(* IEC 61131-3 sources: SemaPLC/sema-plc-benchmark/spec2control-benchmark/data/st-baseline/lng-production/pous/programs, 7 files *)

(* ---- main.st ---- *)
PROGRAM main
VAR
	Heartbeat : bool;
END_VAR

(* Entry point required by OpenPLC Editor v4. The process sections run as parallel program instances under task0; main only provides a scan heartbeat. *)
Heartbeat := NOT Heartbeat;

END_PROGRAM

(* ---- Section2.st ---- *)
PROGRAM Section2
VAR
	FT_101_Flow_PV : real;
	IT_102_Flow_PV : real;
	DP_101_DiffP_PV : real;
	DP_102_DiffP_PV : real;
	LT_101_Level_PV : real;
	IIC_101_LiqSepFlow_SP : real;
	DP_101 : ANALOG_IN;
	DP_102 : ANALOG_IN;
	FT_101 : ANALOG_IN;
	IT_102 : ANALOG_IN;
	LT_101 : ANALOG_IN;
	IIC_101 : RATIO_CONTROL;
	LCV_101 : VALVE_ELECTRIC;
	LCV101_Inhibit_OR : bool;
	IIC101_Inhibit_OR : bool;
END_VAR

DP_101(
    Alarm_Enable := TRUE);
DP_102(
    Alarm_Enable := TRUE);
FT_101(
    Scaling_Slope := 312.5,
    Scaling_Offset := -1250.0,
    Alarm_Enable := TRUE);
IT_102(
    Scaling_Slope := 125.0,
    Scaling_Offset := -500.0,
    Alarm_Enable := TRUE);
LT_101(
    Alarm_Enable := TRUE);
IIC101_Inhibit_OR := LT_101.High_Alarm OR FT_101.Low_Alarm OR DP_101.High_Alarm OR DP_102.High_Alarm;
IIC_101(
    Auto := TRUE,
    PrimaryPV := FT_101.PV,
    SecondaryPV := IT_102.PV,
    RatioSP := 2.5,
    Bias := 0.0,
    MV_MIN := 0.0,
    MV_MAX := 100.0,
    Inhibit := IIC101_Inhibit_OR);
LCV101_Inhibit_OR := FT_101.Low_Alarm OR IT_102.High_Alarm OR IT_102.Low_Alarm OR DP_101.High_Alarm OR DP_102.High_Alarm;
LCV_101(
    Control_Signal := IIC_101.SlaveSP,
    Manual_Mode := FALSE,
    Open_Limit := 100.0,
    Close_Limit := 0.0,
    Inhibit := LCV101_Inhibit_OR);

(* Outputs published to other sections / HMI. *)
FT_101_Flow_PV := FT_101.PV;
IT_102_Flow_PV := IT_102.PV;
DP_101_DiffP_PV := DP_101.PV;
DP_102_DiffP_PV := DP_102.PV;
LT_101_Level_PV := LT_101.PV;
IIC_101_LiqSepFlow_SP := IIC_101.SlaveSP;

END_PROGRAM

(* ---- Section3.st ---- *)
PROGRAM Section3
VAR
	TT201_Temperature_PV : real;
	PT201_FlashTankPressure_PV : real;
	LT201_AbsorberLevel_PV : real;
	AI201_CO2_PV : real;
	TIC201_MV_SteamValveCmd : real;
	AI_201 : ANALOG_IN;
	LT_201 : ANALOG_IN;
	PT_201 : ANALOG_IN;
	TT_201 : ANALOG_IN;
	TIC_201 : PID_BASIC;
	FV_101 : VALVE_ELECTRIC;
	TIC201_Inhibit_OR : bool;
	FV101_Inhibit_OR : bool;
END_VAR

AI_201(
    Alarm_Enable := TRUE);
LT_201(
    Alarm_Enable := TRUE);
PT_201(
    PV_Low := 0.5,
    Alarm_Enable := TRUE);
TT_201(
    PV_High := 50.0,
    Scaling_Slope := 6.25,
    Scaling_Offset := -25.0,
    Alarm_Enable := TRUE);
TIC201_Inhibit_OR := TT_201.High_Alarm OR PT_201.Low_Alarm OR AI_201.High_Alarm OR TT_201.General_Fault;
FV101_Inhibit_OR := TIC201_Inhibit_OR OR LT_201.Low_Alarm;
FV_101(
    Control_Signal := TIC_201.XOUT,
    Manual_Mode := FALSE,
    Open_Limit := 100.0,
    Close_Limit := 0.0,
    Inhibit := FV101_Inhibit_OR);
TIC_201(
    AUTO := TRUE,
    PV := TT_201.PV,
    SP := 45.0,
    MV_MIN := 0.0,
    MV_MAX := 100.0,
    X0 := FV_101.Feedback_Pos,
    KP := 3.0,
    TR := 1.5,
    TD := 0.0,
    Deviation_Limit := 5.0,
    Inhibit := TIC201_Inhibit_OR);

(* Outputs published to other sections / HMI. *)
TT201_Temperature_PV := TT_201.PV;
PT201_FlashTankPressure_PV := PT_201.PV;
LT201_AbsorberLevel_PV := LT_201.PV;
AI201_CO2_PV := AI_201.PV;
TIC201_MV_SteamValveCmd := TIC_201.XOUT;

END_PROGRAM

(* ---- Section4.st ---- *)
PROGRAM Section4
VAR
	AI302_H2O_Outlet_PV : real;
	AI303_Hg_Permissive_PV : real;
	AI304_H2O_RatioOpt_PV : real;
	FT301_FeedGasFlow_PV : real;
	DP301_MolSieveBed_DP_PV : real;
	FFIC303_RegenFlow_SP_to_FIC302 : real;
	AI_302 : ANALOG_IN;
	AI_303 : ANALOG_IN;
	AI_304 : ANALOG_IN;
	DI_301 : DIGITAL_IN;
	DP_301 : ANALOG_IN;
	FIC_302 : PID_BASIC;
	FT_301 : ANALOG_IN;
	FV_302 : VALVE_ELECTRIC;
	FFIC_303 : RATIO_CONTROL;
	Inhibit_OR : bool;
END_VAR

AI_302(
    Alarm_Enable := TRUE);
AI_303(
    Alarm_Enable := TRUE);
AI_304(
    PV_High := 10.0,
    Alarm_Enable := TRUE);
DI_301();
DP_301(
    PV_High := 20.0,
    Alarm_Enable := TRUE);
FT_301(
    PV_Low := 500.0,
    Scaling_Slope := 6.25,
    Scaling_Offset := -25.0,
    Alarm_Enable := TRUE);
Inhibit_OR := AI_302.High_Alarm OR AI_303.High_Alarm OR AI_302.General_Fault OR AI_303.General_Fault OR DI_301.DI_Out OR FT_301.Low_Alarm OR DP_301.High_Alarm;
FFIC_303(
    Auto := TRUE,
    PrimaryPV := FT_301.PV,
    RatioSP := 0.25,
    Bias := 0.0,
    MV_MIN := 0.0,
    MV_MAX := 100.0,
    Inhibit := Inhibit_OR);
FIC_302(
    AUTO := TRUE,
    SP := FFIC_303.SlaveSP,
    MV_MIN := 0.0,
    MV_MAX := 100.0,
    Inhibit := Inhibit_OR);
FV_302(
    Control_Signal := FIC_302.XOUT,
    Open_Limit := 100.0,
    Close_Limit := 0.0,
    Inhibit := Inhibit_OR);

(* Outputs published to other sections / HMI. *)
AI302_H2O_Outlet_PV := AI_302.PV;
AI303_Hg_Permissive_PV := AI_303.PV;
AI304_H2O_RatioOpt_PV := AI_304.PV;
FT301_FeedGasFlow_PV := FT_301.PV;
DP301_MolSieveBed_DP_PV := DP_301.PV;
FFIC303_RegenFlow_SP_to_FIC302 := FFIC_303.SlaveSP;

END_PROGRAM

(* ---- Section5.st ---- *)
PROGRAM Section5
VAR
	PVT_401_Voted_Pressure : real;
	TVT_402_Voted_Temperature : real;
	PT_401A : ANALOG_IN;
	PT_401B : ANALOG_IN;
	PT_401C : ANALOG_IN;
	TT_105 : ANALOG_IN;
	TT_106 : ANALOG_IN;
	TT_107 : ANALOG_IN;
	PVT_401 : VOTING_ANALOG;
	TVT_402 : VOTING_ANALOG;
	PIC_401 : PID_BASIC;
	TIC_402 : PID_BASIC;
	PV_102 : VALVE_ELECTRIC;
	FV_107 : VALVE_ELECTRIC;
	XV_104 : VALVE_ON_OFF;
	I_401 : BOOL_INPUT;
	I_402 : BOOL_INPUT;
	MA_401 : BOOL_INPUT;
	PV102_Inhibit_OR : bool;
	AllPTBad_AND : bool;
	FV107_Inhibit_OR : bool;
	MasterAlarm_OR : bool;
END_VAR

PT_401A(
    PV_High := 2.0,
    PV_Low := 1.6,
    Alarm_Enable := TRUE);
PT_401B(
    PV_High := 2.0,
    PV_Low := 1.6,
    Alarm_Enable := TRUE);
PT_401C(
    PV_High := 2.0,
    PV_Low := 1.6,
    Alarm_Enable := TRUE);
TT_105(
    Alarm_Enable := TRUE);
TT_106(
    Alarm_Enable := TRUE);
TT_107(
    Alarm_Enable := TRUE);
PVT_401(
    Input1 := PT_401A.PV,
    Input2 := PT_401B.PV,
    Input3 := PT_401C.PV,
    Deviation_Limit := 0.09,
    Voting_Scheme := '2oo3',
    EnableAlarm := TRUE);
TVT_402(
    Input1 := TT_105.PV,
    Input2 := TT_106.PV,
    Input3 := TT_107.PV,
    Deviation_Limit := 2.0,
    Voting_Scheme := 'Median',
    EnableAlarm := TRUE);
PIC_401(
    AUTO := TRUE,
    PV := PVT_401.Voted_Output,
    SP := 1.8,
    MV_MIN := 0.0,
    MV_MAX := 100.0);
TIC_402(
    AUTO := TRUE,
    PV := TVT_402.Voted_Output,
    SP := 65.0,
    MV_MIN := 0.0,
    MV_MAX := 100.0);
PV102_Inhibit_OR := PVT_401.Alarm_Voting_Error OR PIC_401.PV_High_Alarm OR PIC_401.PV_Low_Alarm;
I_401(
    Bool_In := PV102_Inhibit_OR,
    Alarm_OnTrue := TRUE,
    Latch_Enable := TRUE);
PV_102(
    Control_Signal := PIC_401.XOUT,
    Open_Limit := 100.0,
    Close_Limit := 0.0,
    Timeout := T#10s,
    Inhibit := I_401.Bool_Out);
FV107_Inhibit_OR := TVT_402.Alarm_Voting_Error OR TIC_402.PV_High_Alarm OR TIC_402.PV_Low_Alarm;
I_402(
    Bool_In := FV107_Inhibit_OR,
    Alarm_OnTrue := TRUE,
    Latch_Enable := TRUE);
FV_107(
    Control_Signal := TIC_402.XOUT,
    Open_Limit := 100.0,
    Close_Limit := 0.0,
    Timeout := T#10s,
    Inhibit := I_402.Bool_Out);
AllPTBad_AND := PT_401A.General_Fault AND PT_401B.General_Fault AND PT_401C.General_Fault;
XV_104(
    Open_Cmd := FALSE,
    Close_Cmd := AllPTBad_AND,
    Timeout := T#5s,
    Inhibit := AllPTBad_AND);
MasterAlarm_OR := PV102_Inhibit_OR OR FV107_Inhibit_OR OR PT_401A.General_Fault OR PT_401B.General_Fault OR PT_401C.General_Fault OR TT_105.General_Fault OR TT_106.General_Fault OR TT_107.General_Fault;
MA_401(
    Bool_In := MasterAlarm_OR,
    Alarm_OnTrue := TRUE,
    Latch_Enable := TRUE);

(* Outputs published to other sections / HMI. *)
PVT_401_Voted_Pressure := PVT_401.Voted_Output;
TVT_402_Voted_Temperature := TVT_402.Voted_Output;

END_PROGRAM

(* ---- Section6.st ---- *)
PROGRAM Section6
VAR
	FT501_PropaneFlow_PV : real;
	FT502_MRFlow_PV : real;
	PT501_EndFlashDrumPressure_PV : real;
	TIT102_MCHE_OutletTemp_PV : real;
	FIC504_MRFlow_SP_From_FFIC503 : real;
	FFIC503_ActiveRatio : real;
	Operator_RatioBias : real;
	FFIC503_DV_HI : bool;
	FFIC503_DV_LO : bool;
	FFIC_503 : RATIO_CONTROL;
	FIC_504 : PID_BASIC;
	FV_502 : VALVE_ELECTRIC;
	FV_501 : VALVE_ELECTRIC;
	FT_501 : ANALOG_IN;
	FT_502 : ANALOG_IN;
	PT_501 : ANALOG_IN;
	TIT_102 : ANALOG_IN;
	FV501_Open_TON : TON;
	RatioDevHi_TON : TON;
	RatioDevLo_TON : TON;
	TempHigh_GT : bool;
	AutoTrim_SEL : real;
	RatioSum_ADD : real;
	RatioBias_ADD : real;
	RatioClamp_LIMIT : real;
	LowFlowCutoff_LT : bool;
	AutoMode_NOT : bool;
	FV501_FullyOpen_GT : bool;
	AutoDisable1_OR : bool;
	AutoDisable3_OR : bool;
	AnySignalIssue_OR : bool;
	ManualSP_SEL1 : real;
	ManualSP_SEL2 : real;
	FT501_RangeAlarm_OR : bool;
	FT502_RangeAlarm_OR : bool;
	FlowRangeViolation_OR : bool;
	FlowSignalFault_OR : bool;
	SafetyCommon_OR : bool;
	RatioDevHi_GT : bool;
	RatioDevLo_LT : bool;
END_VAR

FV_501(
    Open_Limit := 100.0);
FV501_FullyOpen_GT := (FV_501.Feedback_Pos > 99.0);
FV501_Open_TON(
    IN := FV501_FullyOpen_GT,
    PT := T#5s);
FT_501(
    Scaling_Slope := 312.5,
    Scaling_Offset := -1250.0,
    Alarm_Enable := TRUE);
LowFlowCutoff_LT := (FT_501.PV < 500.0);
AutoDisable1_OR := LowFlowCutoff_LT OR FV501_Open_TON.Q;
FT501_RangeAlarm_OR := FT_501.Low_Alarm OR FT_501.High_Alarm;
FT_502(
    Scaling_Slope := 125.0,
    Scaling_Offset := -500.0,
    Alarm_Enable := TRUE);
FT502_RangeAlarm_OR := FT_502.Low_Alarm OR FT_502.High_Alarm;
FlowRangeViolation_OR := FT501_RangeAlarm_OR OR FT502_RangeAlarm_OR;
FlowSignalFault_OR := FT_501.General_Fault OR FT_502.General_Fault;
AnySignalIssue_OR := FlowRangeViolation_OR OR FlowSignalFault_OR;
PT_501(
    Alarm_Enable := TRUE);
SafetyCommon_OR := PT_501.Low_Alarm OR AnySignalIssue_OR;
AutoDisable3_OR := AutoDisable1_OR OR SafetyCommon_OR;
AutoMode_NOT := NOT AutoDisable3_OR;
ManualSP_SEL1 := SEL(G := FV501_Open_TON.Q, IN0 := 100.0, IN1 := 1000.0);
ManualSP_SEL2 := SEL(G := AnySignalIssue_OR, IN0 := ManualSP_SEL1, IN1 := 500.0);
TIT_102(
    PV_High := -155.0,
    Alarm_Enable := TRUE);
TempHigh_GT := (TIT_102.PV > -155.0);
AutoTrim_SEL := SEL(G := TempHigh_GT, IN0 := 0.0, IN1 := 0.1);
RatioSum_ADD := 2.5 + AutoTrim_SEL;
RatioBias_ADD := RatioSum_ADD + Operator_RatioBias;
RatioClamp_LIMIT := LIMIT(MN := 2.0, IN := RatioBias_ADD, MX := 3.0);
FFIC_503(
    Auto := AutoMode_NOT,
    PrimaryPV := FT_501.PV,
    SecondaryPV := FT_502.PV,
    RatioSP := RatioClamp_LIMIT,
    ManOut := ManualSP_SEL2,
    Inhibit := SafetyCommon_OR);
FIC_504(
    PV := FT_502.PV,
    SP := FFIC_503.SlaveSP,
    Inhibit := FlowSignalFault_OR);
FV_502(
    Control_Signal := FIC_504.XOUT);
RatioDevHi_GT := (FFIC_503.RatioErr > 0.2);
RatioDevHi_TON(
    IN := RatioDevHi_GT,
    PT := T#10s);
RatioDevLo_LT := (FFIC_503.RatioErr < -0.2);
RatioDevLo_TON(
    IN := RatioDevLo_LT,
    PT := T#10s);

(* Outputs published to other sections / HMI. *)
FFIC503_DV_HI := RatioDevHi_TON.Q;
FFIC503_DV_LO := RatioDevLo_TON.Q;
FT501_PropaneFlow_PV := FT_501.PV;
FT502_MRFlow_PV := FT_502.PV;
PT501_EndFlashDrumPressure_PV := PT_501.PV;
TIT102_MCHE_OutletTemp_PV := TIT_102.PV;
FIC504_MRFlow_SP_From_FFIC503 := FFIC_503.SlaveSP;
FFIC503_ActiveRatio := FFIC_503.ActiveRatio;

END_PROGRAM

(* ---- Section7.st ---- *)
PROGRAM Section7
VAR
	FT601A_Raw_mA : real;
	FT601B_Raw_mA : real;
	LIT601_Raw_mA : real;
	LT601_Raw_mA : real;
	HS601_HandSwitch_IN : bool;
	FT601A_LNG_Flow_PV : real;
	FT601B_BOG_Flow_PV : real;
	FT601B_BOG_Flow_SP : real;
	LIT601_TankLevel_PV : real;
	LT601_TankLevel_PV : real;
	FT_601A : ANALOG_IN;
	FT_601B : ANALOG_IN;
	LIT_601 : ANALOG_IN;
	LT_601 : ANALOG_IN;
	HS_601 : BOOL_INPUT;
	FFIC_601 : RATIO_CONTROL;
	FIC_601B : PID_BASIC;
	FV_601B : VALVE_ELECTRIC;
	C_601 : MOTOR_ON_OFF;
	RatioControlInhibit : bool;
	CompressorInhibit : bool;
END_VAR

FT_601A(
    Raw_Signal := FT601A_Raw_mA,
    PV_High := 4500.0,
    PV_Low := 100.0,
    Scaling_Slope := 312.5,
    Scaling_Offset := -1250.0,
    Alarm_Enable := TRUE);
FT_601B(
    Raw_Signal := FT601B_Raw_mA,
    PV_High := 900.0,
    PV_Low := 50.0,
    Scaling_Slope := 62.5,
    Scaling_Offset := -250.0,
    Alarm_Enable := TRUE);
LIT_601(
    Raw_Signal := LIT601_Raw_mA,
    Scaling_Slope := 6.25,
    Scaling_Offset := -25.0,
    Alarm_Enable := TRUE);
LT_601(
    Raw_Signal := LT601_Raw_mA,
    Scaling_Slope := 6.25,
    Scaling_Offset := -25.0);
HS_601(
    Bool_In := HS601_HandSwitch_IN,
    Alarm_OnTrue := TRUE);
FIC_601B(
    AUTO := TRUE,
    PV := FT_601B.PV,
    SP := FFIC_601.SlaveSP,
    MV_MIN := 0.0,
    MV_MAX := 100.0,
    X0 := 0.0,
    Deviation_Limit := 100.0,
    Inhibit := LIT_601.High_Alarm);
RatioControlInhibit := HS_601.Alarm_Active OR LIT_601.High_Alarm OR FT_601A.Low_Alarm OR FT_601A.General_Fault OR FT_601B.General_Fault OR FIC_601B.Deviation_Alarm;
FFIC_601(
    Auto := TRUE,
    PrimaryPV := FT_601A.PV,
    SecondaryPV := FT_601B.PV,
    RatioSP := 0.2,
    Bias := 0.0,
    TrimKp := 0.0,
    TrimTi := T#0s,
    MV_MIN := 0.0,
    MV_MAX := 1000.0,
    ManOut := 0.0,
    Inhibit := RatioControlInhibit);
FV_601B(
    Control_Signal := FIC_601B.XOUT,
    Manual_Mode := FALSE,
    Manual_Position := 0.0,
    Open_Limit := 100.0,
    Close_Limit := 0.0,
    Timeout := T#5s,
    Inhibit := LIT_601.High_Alarm);
CompressorInhibit := LIT_601.Low_Alarm OR FV_601B.Alarm OR FT_601A.General_Fault OR FV_601B.Position_Error;
C_601(
    Inhibit := CompressorInhibit);

(* Outputs published to other sections / HMI. *)
FT601A_LNG_Flow_PV := FT_601A.PV;
FT601B_BOG_Flow_PV := FT_601B.PV;
FT601B_BOG_Flow_SP := FFIC_601.SlaveSP;
LIT601_TankLevel_PV := LIT_601.PV;
LT601_TankLevel_PV := LT_601.PV;

END_PROGRAM
